Fanuc KAREL source: ks00038.KL

-- PROVISIONAL review KL for V770-1; original PC SHA256 d271b782dfd7e3fb24af94e9594abcfa4858b0c3408e24b8abd39b3e0532e330
-- Incomplete behavior may be omitted. Consult companion uncertainty JSON. Do not deploy.
PROGRAM KS00038
%NOLOCKGROUP
BEGIN
  -- UNRESOLVED_PC offsets 5-13; opcodes 3F,75
  -- UNRESOLVED_PC offsets 18-27; opcodes 3F,75
  -- UNRESOLVED_PC offsets 32-46; opcodes 22,22,1E
  -- UNRESOLVED_PC offsets 51-55; opcodes 7F
END KS00038
